(* IEC 61131-3 sources: RootPLC/web/playground/examples, 4 files *)

(* ---- 2-star-delta.st ---- *)
(* title: Star-delta motor starter (safety interlock)
   hint: Run plant, then switch start on: star for 5 s, a 100 ms pause, then delta. Test proves star and delta are never on together. *)
FUNCTION_BLOCK FB_StarDelta
VAR_INPUT
    start, stop : BOOL;
END_VAR
VAR_OUTPUT
    main, star, delta : BOOL;
END_VAR
VAR
    st : INT;
    t : TON;
END_VAR
IF stop THEN
    st := 0;
ELSIF start AND st = 0 THEN
    st := 1;
END_IF
CASE st OF
    1:
        t(IN := TRUE, PT := T#5s);
        IF t.Q THEN
            st := 2;
            t(IN := FALSE);
            t(IN := TRUE, PT := T#100ms);
        END_IF
    2:
        t(IN := TRUE, PT := T#100ms);
        IF t.Q THEN
            st := 3;
            t(IN := FALSE);
        END_IF
ELSE
    t(IN := FALSE);
END_CASE
main := st > 0;
star := st = 1;
delta := st = 3;
END_FUNCTION_BLOCK

PROGRAM PRG_StarDelta
VAR_INPUT
    start, stop : BOOL;
END_VAR
VAR_OUTPUT
    main, star, delta : BOOL;
END_VAR
VAR
    sd : FB_StarDelta;
END_VAR
sd(start := start, stop := stop, main => main, star => star, delta => delta);
END_PROGRAM

TEST never_star_and_delta_together
VAR uut : FB_StarDelta; i, both : INT; END_VAR
uut(start := TRUE);
FOR i := 1 TO 700 DO
    uut(start := FALSE);
    IF uut.star AND uut.delta THEN both := both + 1; END_IF
    ADVANCE(T#10ms);
END_FOR
ASSERT_EQ(0, both);
ASSERT_TRUE(uut.delta);
END_TEST

(* ---- 1-traffic-light.st ---- *)
(* title: Traffic light (timers, CASE)
   hint: Press Run plant and switch enable on: green 10 s, yellow 3 s, red 12 s. Press Test to run the TEST block in virtual time. *)
PROGRAM PRG_TrafficLight
VAR_INPUT
    enable : BOOL;
END_VAR
VAR_OUTPUT
    red, yellow, green : BOOL;
END_VAR
VAR
    phase : INT;
    tmr : TON;
    pt : TIME;
    was_enabled : BOOL;
END_VAR
IF NOT enable THEN
    phase := 2;
    tmr(IN := FALSE);
    was_enabled := FALSE;
ELSE
    IF NOT was_enabled THEN
        phase := 0;
        tmr(IN := FALSE);
        was_enabled := TRUE;
    END_IF
    CASE phase OF
        0: pt := T#10s;
        1: pt := T#3s;
    ELSE
        pt := T#12s;
    END_CASE
    tmr(IN := TRUE, PT := pt);
    IF tmr.Q THEN
        phase := (phase + 1) MOD 3;
        CASE phase OF
            0: pt := T#10s;
            1: pt := T#3s;
        ELSE
            pt := T#12s;
        END_CASE
        tmr(IN := FALSE);
        tmr(IN := TRUE, PT := pt);
    END_IF
END_IF
green := enable AND phase = 0;
yellow := enable AND phase = 1;
red := NOT enable OR phase = 2;
END_PROGRAM

TEST cycle_reaches_yellow
VAR uut : PRG_TrafficLight; i : INT; END_VAR
FOR i := 1 TO 115 DO
    uut(enable := TRUE);
    ADVANCE(T#100ms);
END_FOR
uut(enable := TRUE);
ASSERT_TRUE(uut.yellow);
ASSERT_FALSE(uut.red OR uut.green);
END_TEST

(* ---- 3-motor-latch-bug.st ---- *)
(* title: Motor latch with a hidden bug (the test catches it)
   hint: This compiles, but it has a classic precedence bug: AND binds tighter than OR, so stop does not win. Press Test to see it caught, then fix the line to (start OR running) AND NOT stop and test again. *)
PROGRAM PRG_Motor
VAR_INPUT
    start, stop : BOOL;
END_VAR
VAR_OUTPUT
    running : BOOL;
END_VAR
running := start OR running AND NOT stop;
END_PROGRAM

TEST start_latches
VAR uut : PRG_Motor; END_VAR
uut(start := TRUE);
uut(start := FALSE);
ASSERT_TRUE(uut.running);
END_TEST

TEST stop_wins_over_start
VAR uut : PRG_Motor; END_VAR
uut(start := TRUE, stop := TRUE);
ASSERT_FALSE(uut.running);
END_TEST

(* ---- 4-conveyor-interlock.st ---- *)
(* title: Conveyor with emergency stop and guard
   hint: Run plant: switch estop_ok and guard_closed on, then start. Switch estop_ok off: the fault latches until reset. *)
PROGRAM PRG_Conveyor
VAR_INPUT
    start, stop, estop_ok, guard_closed, reset : BOOL;
END_VAR
VAR_OUTPUT
    motor, fault : BOOL;
END_VAR
IF NOT estop_ok THEN
    fault := TRUE;
ELSIF reset THEN
    fault := FALSE;
END_IF
IF fault OR NOT guard_closed OR stop THEN
    motor := FALSE;
ELSIF start THEN
    motor := TRUE;
END_IF
END_PROGRAM

TEST estop_latches_fault
VAR uut : PRG_Conveyor; END_VAR
uut(start := TRUE, estop_ok := TRUE, guard_closed := TRUE);
uut(start := FALSE);
uut(estop_ok := FALSE);
ASSERT_TRUE(uut.fault);
ASSERT_FALSE(uut.motor);
END_TEST
